Fanuc KAREL source: kt00135.KL

-- PROVISIONAL review KL for V770-1; original PC SHA256 24df61125669ed492a371340d805080bb0cb9abe309ad3a8940f3edd87090ba5
-- Incomplete behavior may be omitted. Consult companion uncertainty JSON. Do not deploy.
PROGRAM KT00135
%NOLOCKGROUP
VAR
  I1 : INTEGER
  OUT : INTEGER
-- UNRESOLVED_DECL H2 type=002017
BEGIN
  -- UNRESOLVED_PC offsets 5-16; opcodes 2E,23
  -- UNRESOLVED_PC offsets 21-35; opcodes 2E,22,9D,33,B4
  -- UNRESOLVED_PC offsets 40-62; opcodes 21,22,9D,33,B3,55,23
  -- UNRESOLVED_PC offsets 67-71; opcodes 7F
END KT00135
